PROGRAM FAST
VAR
	(* Enummerations *)

	(* Variables *)

	(* References *)

	(* Interfaces *)

	(* Instances *)

END_VAR


;

END_PROGRAM

(* stored: Version 1.1.0.1, ProductVersion 3.1.4024.15
   POU FAST: Id {66528a3f-d580-4b97-ac35-d6255169dfab}, SpecialFunc None *)
